FUNCTION_BLOCK LongHandshake
VAR_INPUT
	ixStrobIn : BOOL;
END_VAR
VAR_OUTPUT
	oxStrobeOne : BOOL;
	oxStrobeTwo : BOOL;
END_VAR
VAR
END_VAR

END_FUNCTION_BLOCK

(* stored: Version 1.1.0.1, ProductVersion 3.1.4024.12
   POU LongHandshake: Id {e1aaeb54-0808-43ec-b44c-58631c901a70}, SpecialFunc None *)
